// TwinCAT 3 PLC project CcsReceiver
// ProgramVersion: 3.1.4023.0
// libraries:
//   ESO ELT CCS Library, * (ESO)
//   ESO ELT Utility Library, * (ESO)
//   ESO LDC Common Library, * (ESO)
//   ESO LDC Motor Library, * (ESO)
//   ESO LDC Timer Library, * (ESO)
//   Tc2_EtherCAT, * (Beckhoff Automation GmbH)
//   Tc2_Standard, * (Beckhoff Automation GmbH)
//   Tc2_System, * (Beckhoff Automation GmbH)
//   Tc2_Utilities, * (Beckhoff Automation GmbH)
//   Tc3_Module, * (Beckhoff Automation GmbH)
//   VisuDialogs, * (System)
// project tree:
//   / GlobalTextList.TcGTLO, PlcTask.TcTTO, Visualization Manager.TcVMO (not stored)
//   POUs/ MAIN.TcPOU
//   VISUs/ GUI_Drot.TcVIS, GUI_MUDPI_RECEIVER.TcVIS, GUI_TIMER.TcVIS
// real-time tasks:
//   TASK PlcTask: cycle T#10ms, priority 20, ADS port 350
// motion (NC):
//   TASK NC-Task 1 SAF: cycle T#2ms, priority 4, ADS port 501
//   TASK NC-Task 1 SVB: cycle T#10ms, priority 8, ADS port 511
//   AXIS DrotMotor (id 7)
//     General: UnitName=°
//     Dynamic: AccelerationMaximum=100, DecelerationMaximum=100, Acceleration=10.01, Deceleration=10.01, Jerk=28.547
//     Velo: Maximum=6.5
//     TargetPosControl: Range=0.001
//     OtherSettings: AllowMotionCmdToSlave=true
//     encoder EncType=1
//       EncPara: ScaleFactorNumerator=1458, ScaleFactorDenominator=26411000
//         Inc: RefSoftSyncMask=#x0000ffff
//         TimeComp: TimeCompMode=1, EncDelayCycles=4
//     drive DrvType=5
//       Analog: VeloReferenz=7.7, ScaleFactorActTorque=0.1
//       TimeComp: TaskDelayCycles=1
//     controller CtrType=6
//       CtrPara: PriorControlFactor=1
//         PosDiffControl: Range=0.2
//         PID: PosKp=50, VeloKp=0.6, VeloTn=0.08
//         Observer: BandWidth=20
// I/O:
//   DEVICE Device 1 (RT-Ethernet Adapter)
// variable links:
//   CcsReceiver/CcsReceiver Instance <-> NC-Task 1 SAF/Axes/DrotMotor
//     PlcTask Inputs/MAIN.drot.motor.Axis.NcToPlc <-> Outputs/ToPlc
//     PlcTask Outputs/MAIN.drot.motor.Axis.PlcToNc <-> Inputs/FromPlc
//   CcsReceiver/CcsReceiver Instance <-> CcsReceiver/CcsReceiver Instance
//     PlcTask Inputs/MAIN.drot.motor.i_nCouplerState <-> PlcTask Outputs/MAIN.sim_drot.q_nCouplerState
//     PlcTask Inputs/MAIN.drot.motor.switches <-> PlcTask Outputs/MAIN.sim_drot.switches
//   CcsReceiver/CcsReceiver Instance <-> TcCOM Objects/Object1 (TcNtpExternalTimeProvider)
//     PlcTask Inputs/MAIN.fbTimer.i_exNtpConnected <-> Diagnostic/bIsConnected
//     PlcTask Inputs/MAIN.fbTimer.i_exNtpExtOffset <-> Outputs/nSysToExtTimeOffset
//     PlcTask Inputs/MAIN.fbTimer.i_exNtpExtTime <-> Outputs/nExtTime
//     PlcTask Inputs/MAIN.fbTimer.i_exNtpSynchronized <-> Diagnostic/bIsSynchronized
//     PlcTask Inputs/MAIN.fbTimer.i_exNtpSysTime <-> Outputs/nSysTime

CONFIGURATION CcsReceiver
    RESOURCE PLC ON TwinCAT3
        TASK PlcTask(INTERVAL := T#10ms, PRIORITY := 20);
        PROGRAM MAIN WITH PlcTask : MAIN;
    END_RESOURCE
END_CONFIGURATION

// ---- POUs/MAIN.TcPOU
PROGRAM MAIN
VAR
	fbTimer: FB_TIME;
	fbReceiver: FB_CCS_RECEIVER;
	{attribute 'OPC.UA.DA':='1'}
	drot:			FB_MA_DROT;
	{attribute 'OPC.UA.DA':='1'}
	sim_drot:	FB_SIM_MOTOR;
	
	
	
END_VAR

fbTimer();
fbReceiver(refTimeObj := fbTimer);
//
//Devices
//
drot(sName:='DROT', sMotorName:= 'DrotMotor', 
	 in_lrRotation :=fbReceiver.tracking_ccs.north_angle,
	 in_lrPupil := fbReceiver.tracking_ccs.pupil_angle,
	 in_lrParallactic :=fbReceiver.tracking_ccs.pa,
	 nNOVRAM_DevId:=0);
	 
sim_drot(ptrCfg:=ADR(drot.motor.cfg), ptrStat:=ADR(drot.motor.stat));

END_PROGRAM

// ---- VISUs/GUI_Drot.TcVIS
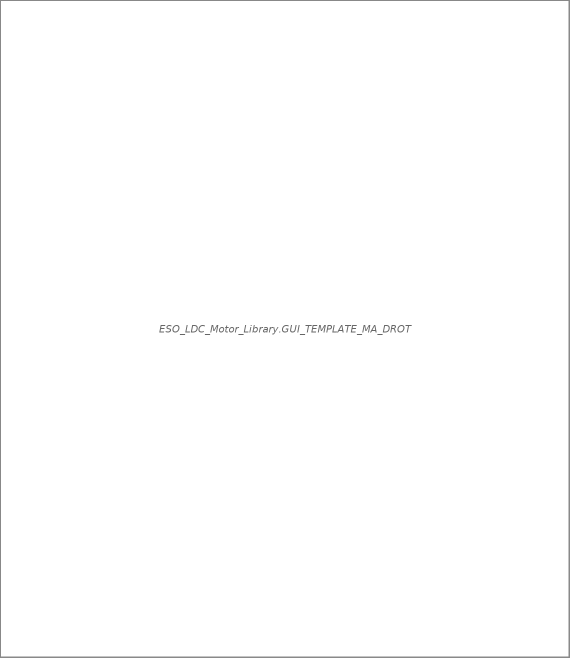
VISUALIZATION GUI_Drot  // 570x658
    Frame (0,0 570x658)
        shows ESO_LDC_Motor_Library.GUI_TEMPLATE_MA_DROT(m_DeviceName := 'drot', m_Instance := MAIN.drot)
END_VISUALIZATION

// ---- VISUs/GUI_MUDPI_RECEIVER.TcVIS
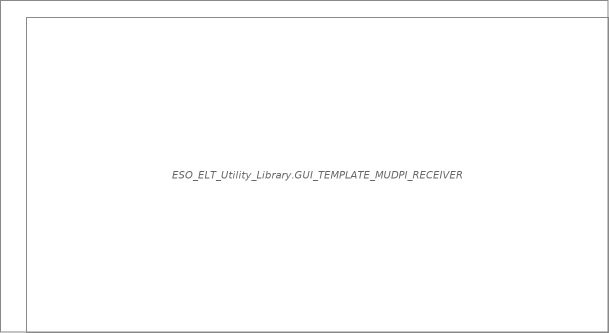
VISUALIZATION GUI_MUDPI_RECEIVER  // 609x333
    Frame (26,17 583x316)
        shows ESO_ELT_Utility_Library.GUI_TEMPLATE_MUDPI_RECEIVER(m_Instance := MAIN.fbReceiver.fbMudpiReceiver)
END_VISUALIZATION

// ---- VISUs/GUI_TIMER.TcVIS
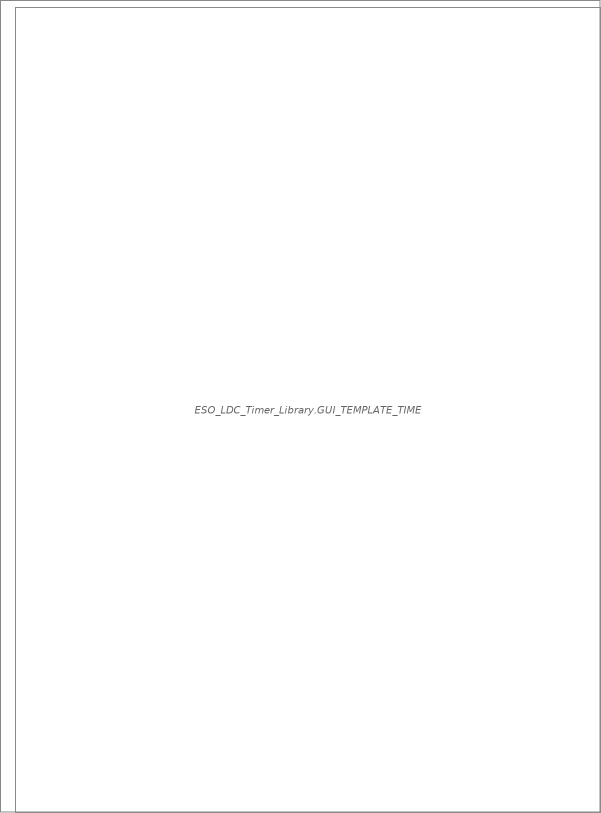
VISUALIZATION GUI_TIMER  // 601x813
    Frame (15,7 586x806)
        shows ESO_LDC_Timer_Library.GUI_TEMPLATE_TIME(m_DeviceName := 'timer', m_Instance := MAIN.fbTimer)
END_VISUALIZATION
